FUNCTION_BLOCK Motor_Generico (* Motor generico (partida direta ou inversor) - HidrycoLib *)
  (* Standard: 61499-2 *)
  (* Version 2.2, 12/11/2026, Hidryco, Hidryco, 2.2: cfgFalhaNA (contato de falha NA). 2.1: velocidade da IHM (STS_VELOCIDADE) em %% entre LSP e HSP lidos do inversor (symlinks stsFrequenciaMaxima HSP 3104, stsFrequenciaMinima LSP 3105); controle continua em Hz. 2.0: inversores ATV600 por Modbus TCP generico (MODBUSGENTCPS unit 248, planilha ATV600 V4.6) no lugar do ATVSpeedControlMbtcp: symlinks com os mesmos nomes em INT (stsVelocidade RFR 0,1 Hz, stsCorrente LCR, stsTensao UOP, stsPotencia OPR, stsTorque OTR, stsCodigoFalha LFT, stsRpm RFRD; stpVelocidade LFR 0,1 Hz; stsFalhaComunicacao = connStatusInt, 1 online), novo cmdPalavraInversor (CMD 8501, bit 7 reset), conversao no basicInversorATV600, cfgEscalaCorrente; com inversor usar cfgSaidaMax = 600 (60,0 Hz = 100 %). 1.9: velocidades da IHM/SCADA em Hz no CLP: STP_SAIDA_MANUAL, STS_VELOCIDADE e STS_VELOCIDADE_REFERENCIA. 1.8: tag STS_FALHA = falha ativa (motor em falha agora, sem memoria). 1.7: alarme de protecao termica sem reconhecimento (ACKTYPE 0) - aparece e some com a termica; velocidade na IHM em Hz (100 % = 60 Hz). 1.6: simbolos sBomba/sMotor/sSoprador - icones de termica e de falha de comunicacao piscam enquanto o alarme nao foi reconhecido. 1.5: symlink stsFalhaComunicacao recebe o ComStatus do ATV (TRUE = comunicacao OK), invertido por NOT para a logica; saida stsComunicacaoOK no CNF. 1.1: padrao SE.App2CommonProcess (supervisao por E_DELAY, horimetro/partidas pelo devMntCalc, escala com limites). 1.3: faceplates ISA-101. 1.4: horimetro com resolucao de 1 s (E_CYCLE + PERSISTENCE), falhas na lista de alarmes do EAE (ALARM_BIT, comunicacao = Warning), reset reconhece os alarmes, termica NF e velocidade manual 50 % por padrao. Campo por symlink ${PATH}: stsFalhaComunicacao, stsRemoto, stsLocal, stsLigado, stsProtecaoTermica, stsSemFalha (NF); saidas cmdAcionamento, stpVelocidade, cmdReset; inversor (cfgInversor=TRUE): stsVelocidade, stsCorrente, stsTensao, stsPotencia, stsFrequencia, stsTorque, stsCodigoFalha, stsRpm *)
  PACKAGE Hidryco.HidrycoLib;
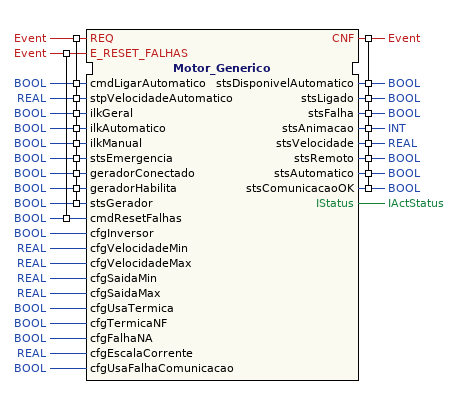
  EVENT_INPUT
    REQ WITH cmdLigarAutomatico, stpVelocidadeAutomatico, ilkGeral, ilkAutomatico, ilkManual, stsEmergencia, geradorConectado, geradorHabilita, stsGerador; (* Atualizacao do processo *)
    E_RESET_FALHAS WITH cmdResetFalhas; (* Reset de falhas pelo processo (com cmdResetFalhas = TRUE) *)
  END_EVENT
  EVENT_OUTPUT
    CNF WITH stsDisponivelAutomatico, stsLigado, stsFalha, stsAnimacao, stsVelocidade, stsRemoto, stsAutomatico, stsComunicacaoOK; (* Status (so na mudanca) *)
  END_EVENT
  VAR_INPUT
    cmdLigarAutomatico : BOOL; (* Comando ligar do processo (modo automatico) *)
    stpVelocidadeAutomatico : REAL; (* Referencia de velocidade do processo (%) *)
    ilkGeral : BOOL; (* Intertravamento geral (automatico e manual) *)
    ilkAutomatico : BOOL; (* Intertravamento so do automatico *)
    ilkManual : BOOL; (* Intertravamento so do manual *)
    stsEmergencia : BOOL; (* Emergencia (TRUE = acionada): retira o comando e exige reset *)
    geradorConectado : BOOL; (* TRUE = o gerador pode alimentar este equipamento *)
    geradorHabilita : BOOL; (* Selecao do operador no CAT Gerador (HAB_GERADOR_EQUIP_n) *)
    stsGerador : BOOL; (* TRUE = planta alimentada pelo gerador *)
    cmdResetFalhas : BOOL; (* Processo: reset de falhas (vale com TRUE) *)
    cfgInversor : BOOL := FALSE; (* TRUE = motor com inversor (referencia de velocidade e medicoes) *)
    cfgVelocidadeMin : REAL := 0.0; (* Limite minimo da referencia de velocidade (%) *)
    cfgVelocidadeMax : REAL := 100.0; (* Limite maximo da referencia de velocidade (%) *)
    cfgSaidaMin : REAL := 0.0; (* Valor de campo equivalente a 0 % (referencia e realimentacao) *)
    cfgSaidaMax : REAL := 100.0; (* Valor de campo equivalente a 100 % (ex.: 100 = %, 60 = Hz, 10000 = Sulzer 0,01 %) *)
    cfgUsaTermica : BOOL := TRUE; (* TRUE = supervisiona a protecao termica *)
    cfgTermicaNF : BOOL := TRUE; (* TRUE = termica NF (FALSE no campo = atuada). Padrao NF (definido pelo usuario) *)
    cfgFalhaNA : BOOL := FALSE; (* TRUE = contato de falha do acionamento NA (TRUE no campo = falha), ligado no symlink stsSemFalha. Padrao FALSE = NF (SEM FALHA) *)
    cfgEscalaCorrente : REAL := 0.1; (* Inversor: A por unidade do LCR (ATV600: 0,1 = LCR em 0,1 A; conferir no display do inversor) *)
    cfgUsaFalhaComunicacao : BOOL := TRUE; (* TRUE = considera o bit de falha de comunicacao da remota *)
  END_VAR
  VAR_OUTPUT
    stsDisponivelAutomatico : BOOL; (* Pode ser comandado pelo automatico agora *)
    stsLigado : BOOL; (* Motor ligado (confirmacao de campo) *)
    stsFalha : BOOL; (* Alguma falha memorizada (exige reset) *)
    stsAnimacao : INT; (* 0 desligado, 1 ligado, 2 falha, 3 manutencao *)
    stsVelocidade : REAL; (* Velocidade real (%); partida direta: 0 ou 100 *)
    stsRemoto : BOOL; (* Chave em remoto *)
    stsAutomatico : BOOL; (* Modo automatico *)
    stsComunicacaoOK : BOOL;
  END_VAR
  PLUGS
    IStatus : IActStatus;
  END_PLUGS
  FBS
    IThis : Motor_Generico_HMI(QI := TRUE);
    plcStart1 : plcStart(Prio := 10);
    Leitura : SYMLINKMULTIVARDST_173DE751D51121F49(QI := TRUE, NAME1 := '$${PATH}stsRemoto', NAME2 := '$${PATH}stsLocal', NAME3 := '$${PATH}stsLigado', NAME4 := '$${PATH}stsProtecaoTermica', NAME5 := '$${PATH}stsSemFalha', NAME6 := '$${PATH}stsFalhaComunicacao'); {SET_ATTRIBUTE(Configuration.GenericFBType.InterfaceParams, Runtime.System#I:=6;VALUE${I$}:BOOL,BOOL,BOOL,BOOL,BOOL,INT)}
    Escrita : SYMLINKMULTIVARSRC_2408DB8E08E99B442(QI := TRUE, NAME1 := '$${PATH}cmdAcionamento', NAME2 := '$${PATH}stpVelocidade', NAME3 := '$${PATH}cmdReset'); {SET_ATTRIBUTE(Configuration.GenericFBType.InterfaceParams, Runtime.System#I:=3;VALUE${I$}:BOOL,INT,BOOL)}
    LeituraInversor1 : SYMLINKMULTIVARDST_15292F208F22048C1(NAME1 := '$${PATH}stsVelocidade', NAME2 := '$${PATH}stsCorrente', NAME3 := '$${PATH}stsTensao', NAME4 := '$${PATH}stsPotencia'); {SET_ATTRIBUTE(Configuration.GenericFBType.InterfaceParams, Runtime.System#I:=4;VALUE${I$}:INT,INT,INT,INT)}
    LeituraInversor2 : SYMLINKMULTIVARDST_15292F208F22048C1(NAME1 := '$${PATH}stsFrequencia', NAME2 := '$${PATH}stsTorque', NAME3 := '$${PATH}stsCodigoFalha', NAME4 := '$${PATH}stsRpm'); {SET_ATTRIBUTE(Configuration.GenericFBType.InterfaceParams, Runtime.System#I:=4;VALUE${I$}:INT,INT,INT,INT)}
    LeituraLimites : SYMLINKMULTIVARDST_184BA62D721027C6E(NAME1 := '$${PATH}stsFrequenciaMaxima', NAME2 := '$${PATH}stsFrequenciaMinima'); {SET_ATTRIBUTE(Configuration.GenericFBType.InterfaceParams, Runtime.System#I:=2;VALUE${I$}:INT,INT)}
    Inversor : basicInversorATV600; (* ATV600 por Modbus generico: brutos -> grandezas; LFR e CMD *)
    EscritaInversor : SYMLINKMULTIVARSRC_5A03F112CD5D470(NAME1 := '$${PATH}cmdPalavraInversor'); {SET_ATTRIBUTE(Configuration.GenericFBType.InterfaceParams, Runtime.System#I:=1;VALUE${I$}:INT)}
    Logica : basicMotorGenerico;
    Supervisao : E_DELAY;
    PulsoReset : E_DELAY(DT := T#3s);
    Tick : E_CYCLE(DT := T#1s);
    PersHorimetro : PERSISTENCE_20652AC5DB8BA8AD5(QI := TRUE); {SET_ATTRIBUTE(Configuration.GenericFBType.InterfaceParams, Runtime.Standard#I:=3;input${I$}:UINT,UINT,UDINT)}
    AlarmeEmergencia : ALARM_BIT(TYPE := 1, ACKTYPE_1 := 2, ACTIVE := TRUE); {SET_ATTRIBUTE(HMI.AlarmText, Emergência acionada)}
    AlarmeTermica : ALARM_BIT(TYPE := 1, ACKTYPE_1 := 0, ACTIVE := TRUE); {SET_ATTRIBUTE(HMI.AlarmText, Proteção térmica atuada)}
    AlarmeAcionamento : ALARM_BIT(TYPE := 1, ACKTYPE_1 := 2, ACTIVE := TRUE); {SET_ATTRIBUTE(HMI.AlarmText, Falha do acionamento (inversor ou soft-starter))}
    AlarmePartida : ALARM_BIT(TYPE := 1, ACKTYPE_1 := 2, ACTIVE := TRUE); {SET_ATTRIBUTE(HMI.AlarmText, Não confirmou a partida no tempo)}
    AlarmeParada : ALARM_BIT(TYPE := 1, ACKTYPE_1 := 2, ACTIVE := TRUE); {SET_ATTRIBUTE(HMI.AlarmText, Não confirmou a parada no tempo)}
    AlarmeComunicacao : ALARM_BIT(TYPE := 1, ACKTYPE_1 := 2, ACTIVE := TRUE); {SET_ATTRIBUTE(HMI.AlarmText, Acionamento sem comunicação)} {SET_ATTRIBUTE(HMI.AlarmClass, Warning)}
    Manutencao : devMntCalc(TBaseOperationDuration := T#1m, TBaseElapsedDuration := T#1d, StateSel := Motor);
    NOT2 : NOT_12669C4E53BA46410; {SET_ATTRIBUTE(Configuration.GenericFBType.InterfaceParams, Runtime.Standard#CNT:=1)}
    E_MERGE1 : E_MERGE;
  END_FBS
  EVENT_CONNECTIONS
    Escrita.INITO TO LeituraLimites.INIT;
    LeituraLimites.CNF TO Inversor.427C31D5944AFC88;
    Leitura.CNF TO Inversor.E4216BCCDF3BB807;
    Inversor.87B3ECE337A4FF70 TO NOT2.REQ;
    LeituraInversor1.CNF TO Inversor.427C31D5944AFC88;
    Inversor.CB0E4FAA64BD8D11 TO Escrita.REQ;
    Inversor.CB0E4FAA64BD8D11 TO EscritaInversor.REQ;
    Escrita.INITO TO EscritaInversor.INIT;
    plcStart1.FIRST_INIT TO IThis.CB1A66AC932C34CE;
    plcStart1.REDO_INIT TO IThis.CB1A66AC932C34CE;
    IThis.60E1F86D6DA4C6BD TO Leitura.INIT;
    Leitura.INITO TO Escrita.INIT;
    Escrita.INITO TO Logica.683CE05B486FAC1D;
    Escrita.INITO TO IThis.EE18699822A64337;
    Escrita.INITO TO Manutencao.INIT;
    Logica.B7169CA02CA38134 TO PersHorimetro.INIT;
    PersHorimetro.INITO TO PersHorimetro.READ;
    PersHorimetro.READCNF TO Logica.84203CA40E4652F0;
    Logica.B3EC08981095182D TO PersHorimetro.WRITE;
    Logica.51A40868F4B890EF TO Tick.START;
    Logica.53ECCF865FC89D5D TO Tick.STOP;
    Tick.EO TO Logica.D2399131CE3E1F66;
    Escrita.INITO TO AlarmeEmergencia.INIT;
    Escrita.INITO TO LeituraInversor1.INIT;
    Escrita.INITO TO LeituraInversor2.INIT;
    REQ TO Logica.5F826E4CBCD659F3;
    REQ TO Logica.9A68BE042B943E25;
    E_RESET_FALHAS TO Logica.0D409FE636F62649;
    Inversor.09B0919BB1BB0E30 TO Logica.9806D419CCC98D7A;
    IThis.EF81D38408160074 TO Logica.079FEC4CDDF030BF;
    IThis.479C30B6853474FB TO Logica.515471E320ACA903;
    IThis.9BF7849A7F6888F9 TO Logica.7C3B0EC5F898F810;
    IThis.E0F935FB34333983 TO Logica.0C2D266AF6549AC9;
    IThis.86D86DF5F3138557 TO Logica.1A33DFD299C36324;
    IThis.D620AE85E607DBF8 TO Manutencao.REQ_RESET;
    Logica.F8CF5B648D94FB56 TO Manutencao.REQ_PV;
    Manutencao.CNF_OPCNT TO Logica.1767A5462AC4396E;
    Logica.78F16FCFC317D932 TO Supervisao.START;
    Logica.551060398A78E95E TO Supervisao.STOP;
    Supervisao.EO TO Logica.F9A311D126CA484B;
    Logica.EEEBF5CC51C91C4E TO PulsoReset.START;
    PulsoReset.EO TO Logica.068D65FB1CCC02E9;
    Logica.0AA258A42CE24B3F TO Inversor.1C34035A3C580B77;
    Logica.D6EF387B8656A6CB TO Inversor.1C34035A3C580B77;
    Logica.78ECC0A7580C66C8 TO E_MERGE1.EI1;
    Logica.78ECC0A7580C66C8 TO IStatus.14377629A1F197A9;
    Logica.0FC40684CDE616F5 TO IStatus.03F1F1C982EE8DD5;
    Logica.0FC40684CDE616F5 TO IStatus.7C93B3F2EA708DB4;
    Logica.814037172F205D14 TO IStatus.BBEA373EFC18FCD4;
    Logica.194428FC25B1C63C TO IThis.102AF7E196740062;
    LeituraInversor2.CNF TO Inversor.427C31D5944AFC88;
    Inversor.09B0919BB1BB0E30 TO IThis.102AF7E196740062;
    AlarmeEmergencia.INITO TO AlarmeEmergencia.REQ_INITDATA;
    AlarmeEmergencia.CNF_INITDATA TO AlarmeEmergencia.ACTIVATE;
    AlarmeEmergencia.INITO TO AlarmeTermica.INIT;
    Logica.194428FC25B1C63C TO AlarmeEmergencia.REQ;
    AlarmeEmergencia.IND_1 TO IThis.102AF7E196740062;
    IThis.E0F935FB34333983 TO AlarmeEmergencia.ACK_C1;
    AlarmeTermica.INITO TO AlarmeTermica.REQ_INITDATA;
    AlarmeTermica.CNF_INITDATA TO AlarmeTermica.ACTIVATE;
    AlarmeTermica.INITO TO AlarmeAcionamento.INIT;
    Logica.194428FC25B1C63C TO AlarmeTermica.REQ;
    AlarmeTermica.IND_1 TO IThis.102AF7E196740062;
    IThis.E0F935FB34333983 TO AlarmeTermica.ACK_C1;
    AlarmeAcionamento.INITO TO AlarmeAcionamento.REQ_INITDATA;
    AlarmeAcionamento.CNF_INITDATA TO AlarmeAcionamento.ACTIVATE;
    AlarmeAcionamento.INITO TO AlarmePartida.INIT;
    Logica.194428FC25B1C63C TO AlarmeAcionamento.REQ;
    AlarmeAcionamento.IND_1 TO IThis.102AF7E196740062;
    IThis.E0F935FB34333983 TO AlarmeAcionamento.ACK_C1;
    AlarmePartida.INITO TO AlarmePartida.REQ_INITDATA;
    AlarmePartida.CNF_INITDATA TO AlarmePartida.ACTIVATE;
    AlarmePartida.INITO TO AlarmeParada.INIT;
    Logica.194428FC25B1C63C TO AlarmePartida.REQ;
    AlarmePartida.IND_1 TO IThis.102AF7E196740062;
    IThis.E0F935FB34333983 TO AlarmePartida.ACK_C1;
    AlarmeParada.INITO TO AlarmeParada.REQ_INITDATA;
    AlarmeParada.CNF_INITDATA TO AlarmeParada.ACTIVATE;
    AlarmeParada.INITO TO AlarmeComunicacao.INIT;
    Logica.194428FC25B1C63C TO AlarmeParada.REQ;
    AlarmeParada.IND_1 TO IThis.102AF7E196740062;
    IThis.E0F935FB34333983 TO AlarmeParada.ACK_C1;
    AlarmeComunicacao.INITO TO AlarmeComunicacao.REQ_INITDATA;
    AlarmeComunicacao.CNF_INITDATA TO AlarmeComunicacao.ACTIVATE;
    AlarmeComunicacao.INITO TO plcStart1.ACK_FIRST;
    Logica.194428FC25B1C63C TO AlarmeComunicacao.REQ;
    AlarmeComunicacao.IND_1 TO IThis.102AF7E196740062;
    IThis.E0F935FB34333983 TO AlarmeComunicacao.ACK_C1;
    NOT2.CNF TO Logica.B2231D0A37008554;
    Leitura.CNF TO E_MERGE1.EI2;
    E_MERGE1.EO TO CNF;
  END_CONNECTIONS
  DATA_CONNECTIONS
    cfgInversor TO LeituraLimites.QI;
    LeituraLimites.VALUE1 TO Inversor.42329CFCD2D17FF4;
    LeituraLimites.VALUE2 TO Inversor.F5C6704A0B387EDE;
    Inversor.AEA206A069529551 TO Logica.3934FBD2505269C1;
    Leitura.VALUE6 TO Inversor.79C0964D27F6F92F;
    Inversor.72B915EBB48AEC2A TO NOT2.IN1;
    LeituraInversor1.VALUE1 TO Inversor.B008AB29C8D9BF35;
    LeituraInversor1.VALUE2 TO Inversor.2D6376362AF121EB;
    LeituraInversor1.VALUE3 TO Inversor.3DFB1C68D576229B;
    LeituraInversor1.VALUE4 TO Inversor.AD5D164EF9FA8C1F;
    LeituraInversor2.VALUE2 TO Inversor.CDF6A5D53E7299DD;
    LeituraInversor2.VALUE3 TO Inversor.292D962FA485B2BC;
    LeituraInversor2.VALUE4 TO Inversor.E045F080AE8FFEBD;
    cfgEscalaCorrente TO Inversor.B66303760760D9ED;
    Logica.6B3311AC79C69555 TO Inversor.2A9BB2F7498BE636;
    Inversor.360DB67778FD2083 TO Escrita.VALUE2;
    Inversor.53A8BE16002FB240 TO EscritaInversor.VALUE1;
    cfgInversor TO EscritaInversor.QI;
    cmdLigarAutomatico TO Logica.193DFCC66FFA3627;
    stpVelocidadeAutomatico TO Logica.98EE3FBBD960BD99;
    ilkGeral TO Logica.32BEE80CEEB8693D;
    ilkAutomatico TO Logica.08FB79476C4E9977;
    ilkManual TO Logica.1B53B44C2D19F3A4;
    geradorConectado TO Logica.08882924EFBEFED3;
    geradorHabilita TO Logica.AFB89A6AEC1EE209;
    cmdResetFalhas TO Logica.1C00AC032E117AF2;
    cfgInversor TO Logica.7320FF5F4A574EDB;
    cfgVelocidadeMin TO Logica.7C3DCCF0844218F0;
    cfgVelocidadeMax TO Logica.E47BA74EEFB23183;
    cfgSaidaMin TO Logica.EDD310DB8258871B;
    cfgSaidaMax TO Logica.B9430F14918E2745;
    cfgUsaTermica TO Logica.28C58F5448A1FB06;
    cfgTermicaNF TO Logica.851269AC75CA9E8E;
    cfgUsaFalhaComunicacao TO Logica.F88C337DE680E3C6;
    stsEmergencia TO Logica.CE80B360618E059C;
    stsGerador TO Logica.C7F3CEE0526BB999;
    cfgInversor TO LeituraInversor1.QI;
    cfgInversor TO LeituraInversor2.QI;
    NOT2.OUT1 TO Logica.14AD61732551E6C9;
    Leitura.VALUE1 TO Logica.4FA04895B58EC5C7;
    Leitura.VALUE2 TO Logica.060151A1F4D195B2;
    Leitura.VALUE3 TO Logica.C82173D2C2DE6C19;
    Leitura.VALUE4 TO Logica.88ACEC8481B97DF2;
    Leitura.VALUE5 TO Logica.6AD75282021BE9C8;
    Inversor.66AEF9F8E70CFE9D TO Logica.D3BA39302C2D6321;
    Logica.689EF5D37ACCCB88 TO Supervisao.DT;
    IThis.503F6CE751BFBAA8 TO Logica.DBE472141CB0338C;
    IThis.8454A63044A9801D TO Logica.E56FE8E891007C74;
    IThis.75974E0F8358E7EE TO Logica.9E5F1B4C72F61C66;
    IThis.947BD655AAF0D307 TO Logica.545E40FBFE122A17;
    IThis.AE42102A3DDDBAD1 TO Logica.6A2A6C1686F090F5;
    IThis.DCF6F7F4874647DD TO Logica.7C364BBDFB8C6BF7;
    IThis.411BDC0B83068DC5 TO Logica.6941FE2305CF8A1E;
    IThis.02D9AF5536125212 TO Manutencao.ResetOperationCount;
    Logica.A2096DD8A524EC3D TO Manutencao.Pv;
    PersHorimetro.output1 TO Logica.3C67B87F17DDB307;
    PersHorimetro.output2 TO Logica.71EDECD1C9B36752;
    PersHorimetro.output3 TO Logica.D6BA299117BFAEF2;
    Logica.750C03D18499F820 TO PersHorimetro.input1;
    Logica.35334824466D36D9 TO PersHorimetro.input2;
    Logica.6F39EF83A6397DAE TO PersHorimetro.input3;
    Manutencao.OperationCount TO Logica.40E1D8559C0FE4D8;
    Logica.FCC70C7B92BB1D0D TO Escrita.VALUE1;
    Logica.0E91B3E8D843667A TO Inversor.B1045E7D3C432FC3;
    Logica.6B3311AC79C69555 TO Escrita.VALUE3;
    Logica.73BD8AC3011DABE5 TO stsDisponivelAutomatico;
    Logica.15F1159202E28B21 TO stsLigado;
    Logica.EBB36D1174CD51D5 TO stsFalha;
    Logica.9E4E2F4C4D54D03D TO stsAnimacao;
    Logica.BEDED4165A410119 TO stsVelocidade;
    Logica.79F308EF21821B91 TO stsRemoto;
    Logica.C042A03D7A6369A4 TO stsAutomatico;
    Logica.79F308EF21821B91 TO IThis.294C3F7487077BBC;
    Logica.A3458504BF6DF144 TO IThis.47A58C942EA6825F;
    Logica.9558D049DB2CB76C TO IThis.45C161DD8A14A557;
    Logica.15F1159202E28B21 TO IThis.3E8EAAE5C56CE832;
    Logica.C042A03D7A6369A4 TO IThis.35FB3D0DD77469AD;
    Logica.608D1BE3AF5D2E15 TO IThis.99D45055626342AC;
    Logica.9E4E2F4C4D54D03D TO IThis.5F2DFD1D3F9171CC;
    Logica.170EA16E9186BAB7 TO IThis.8C20ADCFDB9510BA;
    Logica.7A11796B672969B4 TO IThis.F05387CCA913E498;
    Logica.7A1632E7C1C3C53A TO IThis.914AB4D395F40992;
    Logica.F8277369617C4FEC TO IThis.F4A10448D767AD4A;
    Logica.24D167508AB5B3BF TO IThis.E3B83D77D62F143A;
    Logica.F939957499D9DE01 TO IThis.67A853C96706FC71;
    Logica.8DBC1E391953B77A TO IThis.05D22B39A9C68F81;
    Logica.47CFEB602576FDE6 TO IThis.F3A94F346E1F2344;
    Logica.524B369F0AC1FCF0 TO IThis.8DFE7C65FD4D26BA;
    Logica.85F7CA319643FCE9 TO IThis.04BB4F9CD24381F2;
    Logica.73BD8AC3011DABE5 TO IThis.21C1E76BA48924FC;
    Logica.6F39EF83A6397DAE TO IThis.16651CA122A2B95B;
    Logica.35334824466D36D9 TO IThis.9D04D7BAE7D40E02;
    Logica.CA7BD048A830149F TO IThis.D7DA16EAB6FF6EEE;
    Logica.F6C8BE93FC698E3B TO IThis.1CEAC095F858B414;
    Logica.B328ACD14E28750E TO IThis.C238ADA8DCED3CBD;
    Logica.E8C96E839FCF2B87 TO IThis.869F2DEDF63D520E;
    AlarmeEmergencia.STATE_1 TO IThis.51C58C818B781512;
    AlarmeTermica.STATE_1 TO IThis.4CD0EDFE6E941B41;
    AlarmeAcionamento.STATE_1 TO IThis.B155B2692776CD13;
    AlarmePartida.STATE_1 TO IThis.7A43BEA87F2F44B9;
    AlarmeParada.STATE_1 TO IThis.EC0AD5583DFA829A;
    AlarmeComunicacao.STATE_1 TO IThis.C1CC4C6B5FCBBCD2;
    Inversor.37526A7D778B9E7B TO IThis.7E0C670138DD7B76;
    Inversor.930BAE86F242A833 TO IThis.6875B6D16C69A2E9;
    Inversor.2DDD2CDD0C674D43 TO IThis.62A08FAA4AB91A15;
    Inversor.2C7FE4FF8CF8442A TO IThis.803D206AACB27DD7;
    Inversor.20BE98C14B2600D9 TO IThis.11AE970559C4D02C;
    Inversor.59458D47837A2DDA TO IThis.A48E8BCAD9763E7A;
    Inversor.49A95C3D64F24BED TO IThis.3ABB296BCC446C60;
    Logica.47CFEB602576FDE6 TO AlarmeEmergencia.INP;
    Logica.F8277369617C4FEC TO AlarmeTermica.INP;
    Logica.24D167508AB5B3BF TO AlarmeAcionamento.INP;
    Logica.F939957499D9DE01 TO AlarmePartida.INP;
    Logica.8DBC1E391953B77A TO AlarmeParada.INP;
    Logica.7A1632E7C1C3C53A TO AlarmeComunicacao.INP;
    Logica.73BD8AC3011DABE5 TO IStatus.9E0B44559326BEAF;
    Logica.15F1159202E28B21 TO IStatus.D41A46B14EF7208D;
    Logica.C9FFC4D7ACE51BE3 TO IStatus.227987A2F0C6A825;
    Logica.BEDED4165A410119 TO IStatus.B9E42D72CEF16844;
    Logica.BEDED4165A410119 TO IStatus.63F2604DAA7CFD9F;
    Logica.D50BA6FDF5BB251B TO IStatus.6786798CC8B69406;
    Inversor.72B915EBB48AEC2A TO stsComunicacaoOK;
    Logica.E6802855A03CB240 TO IThis.43C738994B732921;
    Logica.5355A350F226F825 TO IThis.06277D222F5F3621;
    Logica.E6B78B01125D043A TO IThis.7B3A3676FBDE5F7A;
    cfgFalhaNA TO Logica.BC9C4A0B25009270;
  END_CONNECTIONS
END_FUNCTION_BLOCK
